(* Logix 5000 project; controller CIP_14485201 vendor 1 type 14 code 216 rev 38.11; software revision 38.01; part 12 of 12 *)
(* tags used below, declared in another part *)
   PID2 : PID;   // SUPPLY FLOW PID
   SCLD_Supply_Flow : SCALE;   // SUPPLY FLOW 0-60 GPM

PROGRAM PID_SupplyFlow   (* main routine _02_SUB *)

ROUTINE _02_SUB   (* ladder *)
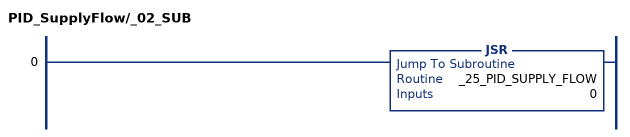
   0: JSR(_25_PID_SUPPLY_FLOW,0);
END_ROUTINE

ROUTINE _25_PID_SUPPLY_FLOW   (* ladder *)
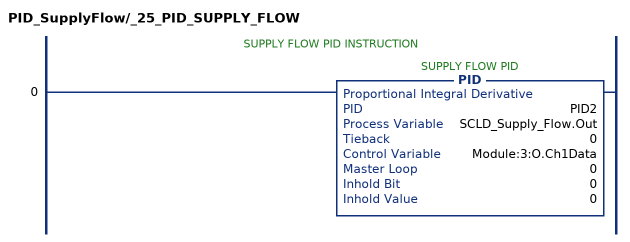
   // SUPPLY FLOW PID INSTRUCTION
   0: PID(PID2,SCLD_Supply_Flow.Out,0,Module:3:O.Ch1Data,0,0,0);
END_ROUTINE
END_PROGRAM
